// TIA Portal V20 export
ORGANIZATION_BLOCK "T7_OB20"   // OB20, LAD, TimeDelayInterrupt
TITLE = T7_OB20
{ S7_Optimized_Access := 'TRUE' }
AUTHOR : IA
FAMILY : PRUEBA
VERSION : 0.1
// Tanda 3: TimeDelayInterrupt, incrementa OB20_Cuenta
// stored: AutoNumber false, IsIECCheckEnabled false, SetENOAutomatically false
   VAR_INPUT
      Sign : Word;
   END_VAR
BEGIN

REGION Network 1: Contador de vida
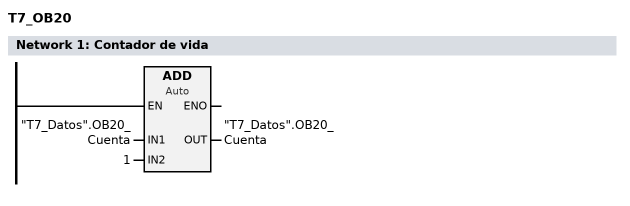
   RUNG wire#powerrail
      Add(in1 := "T7_Datos".OB20_Cuenta, in2 := 1, out => "T7_Datos".OB20_Cuenta)
   END_RUNG
   // the same network as SCL:
   "T7_Datos".OB20_Cuenta := "T7_Datos".OB20_Cuenta + 1;
END_REGION
END_ORGANIZATION_BLOCK
